// TIA Portal V21 export
// export: Created 2026-10-24T00:39:25.7362804Z, ExportSetting WithDefaults, DisplayName Totally Integrated Automation Portal, DisplayVersion V21 Update 1, DisplayName SINAMICS Startdrive Advanced, DisplayVersion V21 HF2, DisplayName SINAMICS Startdrive G110M, G120, G120C, G120D, G120P, G115D, DisplayVersion V21 HF2, DisplayName SINAMICS Startdrive G130, G150, S120, S150, G200, G220, S200, S210, S220, Innomotics MVD, DisplayVersion V21 HF2, DisplayName STEP 7 Professional, DisplayVersion V21 Update 1, DisplayName STEP 7 Safety, DisplayVersion V21, DisplayName Tech WebApplication, DisplayVersion V21, DisplayName WinCC Basic/Comfort/Advanced, DisplayVersion V21 Update 1, DisplayName WinCC Unified, DisplayVersion V21 Update 1
VAR_GLOBAL   // PLC tag table "Tags_Openness"
   OpnStart AT %I4.0 : Bool;   // Start input, exported through Openness
   OpnFlow AT %IW6 : Word;   // Raw flow
   OpnLamp AT %Q4.0 : Bool;   // Lamp output
   OpnHelper AT %M20.0 : Bool;   // Helper bit
   OpnHidden AT %MW22 : Int;   // Not accessible from HMI   {ExternalVisible false, ExternalWritable false}
END_VAR
VAR_GLOBAL CONSTANT   // user constants
   OPN_LIMIT : Int := 250;   // Upper limit
END_VAR
